FUNCTION_BLOCK ResetConfSemIlck (* ConfResetReq efetivo: ConfResetIn AND NOT SemReset (alarme de realimentacao nao pede reset na janela de intertravamento) *)
  (* Standard: 61499-2 *)
  (* Version 1.1, 05/11/2026, Hidryco, Hidryco, 1.1: eventos de saida listados no ECAction (sem isso o runtime nao emite nenhum; o ST so liga/desliga). 1.0: ConfResetOut = ConfResetIn AND NOT SemReset; repassa o REQ (gera CNF sempre) para o REQ_PARA do controle. *)
  PACKAGE SE.Nereda;
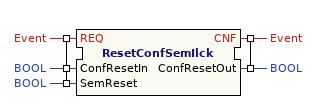
  EVENT_INPUT
    REQ WITH ConfResetIn, SemReset; (* Parametros ou janela mudaram *)
  END_EVENT
  EVENT_OUTPUT
    CNF WITH ConfResetOut; (* Para o REQ_PARA do controle *)
  END_EVENT
  VAR_INPUT
    ConfResetIn : BOOL; (* ConfResetReq da IHM *)
    SemReset : BOOL; (* Janela de intertravamento *)
  END_VAR
  VAR_OUTPUT
    ConfResetOut : BOOL; (* ConfResetReq para o controle *)
  END_VAR
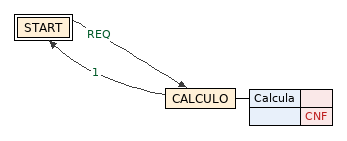
  EC_STATES
    START; (* Estado inicial *)
    CALCULO : Calcula, -> CNF; (* Calcula; o algoritmo decide quais eventos saem *)
  END_STATES
  EC_TRANSITIONS
    START TO CALCULO := REQ;
    CALCULO TO START := 1;
  END_TRANSITIONS
  ALGORITHM Calcula IN ST: (* ConfResetReq efetivo: ConfResetIn AND NOT SemReset (alarme de realimentacao nao pede reset na janela de intertravamento) *)
ConfResetOut := ConfResetIn AND NOT SemReset;
CNF := TRUE;
  END_ALGORITHM
END_FUNCTION_BLOCK
